{region 'Documentation'}
(*!
<summary>Checks that selected bits match the expected masked value.</summary>
*)
{endregion}
FUNCTION_BLOCK AssertEqualMask_Word EXTENDS AssertionBase
VAR_INPUT
    IN : WORD; //! Actual bitfield.
    Mask : WORD := 16#FFFF; //! Selects evaluated bits; defaults to all bits. An empty mask produces Error during evaluation.
    Expected : WORD; //! Expected value; bits outside Mask are ignored.
END_VAR

SUPER^();

{region 'Documentation'}
(*!
<summary>Rejects an empty mask before comparing selected bits.</summary>
*)
{endregion}
METHOD PROTECTED Assert
VAR
    Message : STRING(GVL_Constants.MessageLength);
    MaskText : STRING(GVL_Constants.AssertionValueLength);
    ExpectedText : STRING(GVL_Constants.AssertionValueLength);
    ActualText : STRING(GVL_Constants.AssertionValueLength);
END_VAR
VAR CONSTANT
    NoMask : WORD := 16#00;
    HexDigitCount : USINT := 4;
END_VAR
IF NOT EvaluationActive THEN
    RETURN;
END_IF;

IF Result = E_Result.Error THEN
    RETURN;
END_IF;

IF Mask = NoMask THEN
    MaskText := CreateAssertionTextValue_Hex(Value := WORD_TO_LWORD(Mask),
        DigitCount := HexDigitCount);
    Message := CONCAT('Assertion error: mask must not be empty. Mask = ',
        MaskText);
    Message := CONCAT(Message, '.');
    Error(Message := Message);
    RETURN;
END_IF;

IF Result = E_Result.Failed THEN
    RETURN;
END_IF;

IF (IN AND Mask) <> (Expected AND Mask) THEN
    MaskText := CreateAssertionTextValue_Hex(Value := WORD_TO_LWORD(Mask),
        DigitCount := HexDigitCount);
    ExpectedText := CreateAssertionTextValue_Hex(Value := WORD_TO_LWORD(Expected),
        DigitCount := HexDigitCount);
    ActualText := CreateAssertionTextValue_Hex(Value := WORD_TO_LWORD(IN),
        DigitCount := HexDigitCount);
    Message := CONCAT('Assertion failed: selected bits do not match. Expected = ',
        ExpectedText);
    Message := CONCAT(Message, ', Mask = ');
    Message := CONCAT(Message, MaskText);
    Message := CONCAT(Message, ', Actual = ');
    Message := CONCAT(Message, ActualText);
    Message := CONCAT(Message, '.');
    Fail(Message := Message);
    RETURN;
END_IF;

Pass();
END_METHOD

END_FUNCTION_BLOCK

(* stored: Version 1.1.0.1
   POU AssertEqualMask_Word: Id {52ac2086-baf9-4189-b043-30a25aec269e}, SpecialFunc None
   Folder Internal: Id {725ea3a2-6160-4c37-8e1a-9782aabf85fc}
   Method Assert: Id {df6bd827-ca58-4325-9389-40626d63f539} *)
